TYPE ST_Bits :
STRUCT
	Bit1:BIT;
	Bit2:BIT;
	Bit3:BIT;
	Bit4:BIT;
	Bit5:BIT;
	Bit6:BIT;
	Bit7:BIT;
	Bit8:BIT;
	Bit9:BIT;
	Bit10:BIT;
	Bit11:BIT;
	Bit12:BIT;
	Bit13:BIT;
	Bit14:BIT;
	Bit15:BIT;
	Bit16:BIT;
END_STRUCT
END_TYPE

(* stored: Version 1.1.0.1
   DUT ST_Bits: Id {10b53587-2221-4ad2-820d-04ebbbb46002} *)
